// TIA Portal V20 export
// export: Created 2026-10-12T05:00:30.3907159Z, ExportSetting WithDefaults, DisplayName Totally Integrated Automation Portal, DisplayVersion V20, DisplayName TIA Portal Openness, DisplayVersion V20, DisplayName TIA Portal Teamcenter Gateway, DisplayVersion V20, DisplayName TIA Portal Version Control Interface, DisplayVersion V20, DisplayName SINAMICS Startdrive Advanced, DisplayVersion V20 SP1 Update 2, DisplayName SINAMICS Startdrive G110M, G120, G120C, G120D, G120P, G115D, DisplayVersion V20 SP1 Update 2, DisplayName SINAMICS Startdrive G130, G150, S120, S150, SINAMICS MV, G220, S200, S210, DisplayVersion V20 SP1 Update 2, DisplayName STEP 7 Professional, DisplayVersion V20, DisplayName STEP 7 Safety, DisplayVersion V20, DisplayName WinCC Basic/Comfort/Advanced, DisplayVersion V20, DisplayName WinCC Professional, DisplayVersion V20, DisplayName WinCC Unified, DisplayVersion V20
FUNCTION "FRK_JsonHeader" : Bool   // FC119, SCL
{ S7_Optimized_Access := 'TRUE' }
VERSION : 0.1
// stored: AutoNumber true, IsIECCheckEnabled false, SetENOAutomatically false, UDAEnableTagReadback false
   VAR_INPUT
      Data : "ST_ConfigSetInfo";
   END_VAR
   VAR_IN_OUT
      Line : WString;
   END_VAR
   VAR_TEMP
      Ok : Bool;
      Flag : WString[1];
   END_VAR
BEGIN

   #FRK_JsonHeader := FALSE;
   #Line := WSTRING#'{';
   #Ok := "FRK_JsonAdd"(Key := 'set', Value := STRING_TO_WSTRING(#Data.SetName), Quoted := TRUE, LastField := FALSE, Line := #Line);
   IF NOT #Ok THEN
       #Line := WSTRING#'';
       RETURN;
   END_IF;
   #Ok := "FRK_JsonAdd"(Key := 'root', Value := STRING_TO_WSTRING(#Data.RootIdentity), Quoted := TRUE, LastField := FALSE, Line := #Line);
   IF NOT #Ok THEN
       #Line := WSTRING#'';
       RETURN;
   END_IF;
   #Ok := "FRK_JsonAdd"(Key := 'schema', Value := UINT_TO_WSTRING(#Data.SetSchema), Quoted := FALSE, LastField := FALSE, Line := #Line);
   IF NOT #Ok THEN
       #Line := WSTRING#'';
       RETURN;
   END_IF;
   #Ok := "FRK_JsonAdd"(Key := 'configRev', Value := UDINT_TO_WSTRING(#Data.ConfigRev), Quoted := FALSE, LastField := FALSE, Line := #Line);
   IF NOT #Ok THEN
       #Line := WSTRING#'';
       RETURN;
   END_IF;
   #Ok := "FRK_JsonAdd"(Key := 'kind', Value := DINT_TO_WSTRING(#Data.Kind), Quoted := FALSE, LastField := FALSE, Line := #Line);
   IF NOT #Ok THEN
       #Line := WSTRING#'';
       RETURN;
   END_IF;
   #Ok := "FRK_JsonAdd"(Key := 'model', Value := STRING_TO_WSTRING(#Data.ModelCode), Quoted := TRUE, LastField := FALSE, Line := #Line);
   IF NOT #Ok THEN
       #Line := WSTRING#'';
       RETURN;
   END_IF;
   #Ok := "FRK_JsonAdd"(Key := 'records', Value := DINT_TO_WSTRING(#Data.RecordCount), Quoted := FALSE, LastField := FALSE, Line := #Line);
   IF NOT #Ok THEN
       #Line := WSTRING#'';
       RETURN;
   END_IF;
   #Ok := "FRK_JsonAdd"(Key := 'created', Value := ULINT_TO_WSTRING(LDT_TO_ULINT(#Data.CreatedAt) / ULINT#1000000000), Quoted := FALSE, LastField := FALSE, Line := #Line);
   IF NOT #Ok THEN
       #Line := WSTRING#'';
       RETURN;
   END_IF;
   IF #Data.TimeSynchronized THEN
       #Flag := WSTRING#'1';
   ELSE
       #Flag := WSTRING#'0';
   END_IF;
   #Ok := "FRK_JsonAdd"(Key := 'clock', Value := #Flag, Quoted := FALSE, LastField := TRUE, Line := #Line);
   IF NOT #Ok THEN
       #Line := WSTRING#'';
       RETURN;
   END_IF;
   #FRK_JsonHeader := TRUE;
END_FUNCTION
